FUNCTION_BLOCK FB_Batch
VAR
    bStart, bAbort, bValveOpen, bLevel : BOOL;
    rTemp : REAL;
    fbMixer : FB_Mixer;
END_VAR

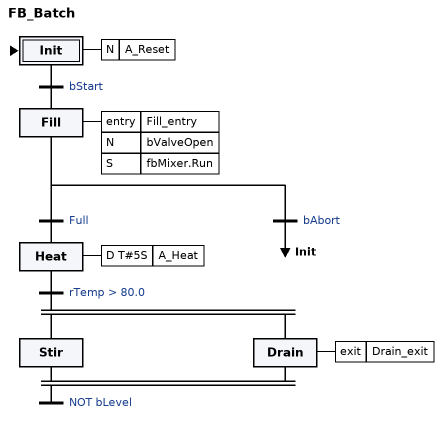
INITIAL_STEP Init:
    A_Reset(N);
END_STEP
TRANSITION FROM Init TO Fill
    := bStart;
END_TRANSITION
STEP Fill:
    Fill_entry(P1);  // entry action
    bValveOpen(N);
    fbMixer.Run(S);
END_STEP
TRANSITION FROM Fill TO Heat
    := Full;
END_TRANSITION
STEP Heat:
    A_Heat(D, T#5S);
END_STEP
TRANSITION FROM Fill TO Init
    := bAbort;
END_TRANSITION
TRANSITION FROM Heat TO (Stir, Drain)
    := rTemp > 80.0;
END_TRANSITION
STEP Stir:
END_STEP
STEP Drain:
    Drain_exit(P0);  // exit action
END_STEP
TRANSITION FROM (Stir, Drain) TO ???
    := NOT bLevel;
END_TRANSITION

ACTION A_Reset:
bValveOpen := FALSE;
END_ACTION

ACTION A_Heat:
rTemp := rTemp + 0.5;
END_ACTION

ACTION Fill_entry:
bLevel := FALSE;
END_ACTION

ACTION Drain_exit:
bValveOpen := FALSE;
END_ACTION

TRANSITION Full:
bLevel AND NOT bAbort
END_TRANSITION

END_FUNCTION_BLOCK

(* stored: Version 1.1.0.1, ProductVersion 3.1.4024.12
   POU FB_Batch: Id {00000000-0000-0000-0000-000000000001}, SpecialFunc None
   Action A_Reset: Id {00000000-0000-0000-0000-000000000011}
   Action A_Heat: Id {00000000-0000-0000-0000-000000000012}
   Action Fill_entry: Id {00000000-0000-0000-0000-000000000013}
   Action Drain_exit: Id {00000000-0000-0000-0000-000000000014}
   Transition Full: Id {00000000-0000-0000-0000-000000000015} *)
